// TIA Portal V20 export
FUNCTION_BLOCK "CONTROL_LINE"   // FB7, LAD
{ S7_Optimized_Access := 'TRUE' }
// stored: MemoryReserve 100, SetENOAutomatically false
   VAR
      TIMER_reset { S7_SetPoint := 'True'} : TON_TIME;
      P_TRIG_INICIAL : Bool;
      P_TRIG_RESET : Bool;
      AUTOMAT { S7_SetPoint := 'True'} : "SENSOR";
      MANUAL { S7_SetPoint := 'True'} : "SENSOR";
      SENSOR_3 { S7_SetPoint := 'True'} : "SENSOR";
      SENSOR_4 { S7_SetPoint := 'True'} : "SENSOR";
      SENSOR_5 { S7_SetPoint := 'True'} : "SENSOR";
      SENSOR_6 { S7_SetPoint := 'True'} : "SENSOR";
      SENSOR_7 { S7_SetPoint := 'True'} : "SENSOR";
      SENSOR_8 { S7_SetPoint := 'True'} : "SENSOR";
      SENSOR_9 { S7_SetPoint := 'True'} : "SENSOR";
      SENSOR_10 { S7_SetPoint := 'True'} : "SENSOR";
      SENSOR_11 { S7_SetPoint := 'True'} : "SENSOR";
      dvere_L_A { S7_SetPoint := 'True'} : "SENSOR";
      dvere_L_B { S7_SetPoint := 'True'} : "SENSOR";
      dvere_P_A { S7_SetPoint := 'True'} : "SENSOR";
      dvere_P_B { S7_SetPoint := 'True'} : "SENSOR";
      SEN_STRUCT : Struct
         AUTOMAT : Bool;
         AUTOMAT_NEG : Bool;
         MANUAL : Bool;
         MANUAL_NEG : Bool;
         SENSOR_TLAKU : Bool;
         SENSOR_TLAKU_NEG : Bool;
         power : Bool;
         power_neg : Bool;
         safety : Bool;
         safety_neg : Bool;
         s_10 : Bool;
         TLA_STOP : Bool;
         TLA_STOP_NEG : Bool;
         TLA_START : Bool;
         TLA_START_NEG : Bool;
         TLA_KVIT : Bool;
         TLA_KVIT_NEG : Bool;
         s_17 : Bool;
         S19 : Bool;
         L1_OK : Bool;
         L1_NOT_OK : Bool;
         L2_OK : Bool;
         L2_NOT_OK : Bool;
         L3_OK : Bool;
         L3_NOT_OK : Bool;
         dvere_L_A : Bool;
         dvere_L_B : Bool;
         dvere_P_A : Bool;
         dvere_P_B : Bool;
         S30 : Bool;
         S31 : Bool;
         LASER_MEMOR : Bool;
      END_STRUCT;
      "M" : Struct
         P_TRIK_hmi_manual : Bool;
         p_trig_hmi_automat : Bool;
         N_TRIG_REZIM : Bool;
         M_4 : Bool;
         hlaseni_chyby : Bool;
         M_6 : Bool;
         M_7 : Bool;
         M_8 : Bool;
         M_9 : Bool;
         p_Trig_al : Bool;
         n_trig_al : Bool;
         p_trig_wro : Bool;
         n_trig_wro : Bool;
         M_14 : Bool;
         M_15 : Bool;
         N_TRIG_MANUAL : Bool;
         M_17 : Bool;
         M_18 : Bool;
         M_19 : Bool;
         M_20 : Bool;
         M_21 : Bool;
         M_22 : Bool;
         M_23 : Bool;
         M_24 : Bool;
         M_25 : Bool;
         M_26 : Bool;
         M_27 : Bool;
         M_28 : Bool;
         M_29 : Bool;
         M_30 : Bool;
         M_31 : Bool;
         M_32 : Bool;
      END_STRUCT;
      trig : Struct
         reset_error_all : Bool;
         TRIG_FOR_OP_4_AUTOMAT : Bool;
         t_3 : Bool;
         t_4 : Bool;
         t_5 : Bool;
         t_6 : Bool;
         t_7 : Bool;
         t_8 : Bool;
      END_STRUCT;
      SQCR : Int;
      job_mailbox : Array[0..3] of Word;
      n_trig_res_auit : Bool;
      inicial_control { S7_SetPoint := 'True'} : TON_TIME;
      SQCR_SAFETY { S7_SetPoint := 'True'} : Int;
      n_trig_RESET_AUT : Bool;
      P_TRIG_RESET_SAFETY : Bool;
      air { S7_SetPoint := 'True'} : TON_TIME;
      HMI_ALARM { S7_SetPoint := 'True'} : Int;
   END_VAR
   VAR_TEMP
      "string" : String;
      smaz_me : Bool;
      majak_green_s1 : Bool;
      majak_red_s1 : Bool;
      majak_yelou_s1 : Bool;
      majak_blue_s1 : Bool;
      majak_orange_s1 : Bool;
      majak_green_s2 : Bool;
      majak_red_s2 : Bool;
      majak_yelou_s2 : Bool;
      majak_blue_s2 : Bool;
      majak_orange_s2 : Bool;
      majak_green_s3 : Bool;
      majak_red_s3 : Bool;
      majak_yelou_s3 : Bool;
      majak_blue_s3 : Bool;
      majak_orange_s3 : Bool;
      majak_green_s4 : Bool;
      majak_red_s4 : Bool;
      majak_yelou_s4 : Bool;
      majak_blue_s4 : Bool;
      majak_orange_s4 : Bool;
      majak_green_s5 : Bool;
      majak_red_s5 : Bool;
      majak_yelou_s5 : Bool;
      majak_blue_s5 : Bool;
      majak_orange_s5 : Bool;
   END_VAR
   VAR CONSTANT
      STEP_0_FIRST_START : Int := 0;
      STEP_3 : Int := 3;
      STEP_5 : Int := 5;
      STEP_10 : Int := 10;
      STEP_15 : Int := 15;
      STEP_20 : Int := 20;
      STEP_25 : Int := 25;
      STEP_27 : Int := 27;
      STEP_30 : Int := 30;
      STEP_35 : Int := 35;
      STEP_40 : Int := 40;
      STEP_45 : Int := 45;
      STEP_48 : Int := 48;
      STEP_50 : Int := 50;
      STEP_52 : Int := 52;
      STEP_55 : Int := 55;
      STEP_60 : Int := 60;
      STEP_65 : Int := 65;
      STEP_70 : Int := 70;
      STEP_75 : Int := 75;
      STEP_80 : Int := 80;
      STEP_85 : Int := 85;
      STEP_90 : Int := 90;
      STEP_95 : Int := 95;
      STEP_100 : Int := 100;
      STEO_105 : Int := 105;
   END_VAR
   VAR_TEMP   // added for the SCL form of the ladder/FBD networks
      _w1 : Bool;
      _w2 : Bool;
      _w3 : Bool;
      _w4 : Bool;
      _w5 : Bool;
   END_VAR
BEGIN

REGION Network 1 (SCL)
   // SET  BASIC ELEMENTS
   // odpojení nepoužívaných kontaktů
   "LOG_0" := 0;
   "LOG_1" := 1;
   "SMAZ_ME_0" := 0;
   "SMAZ_ME_1" := 1;
END_REGION

REGION Network 2: SENSORS
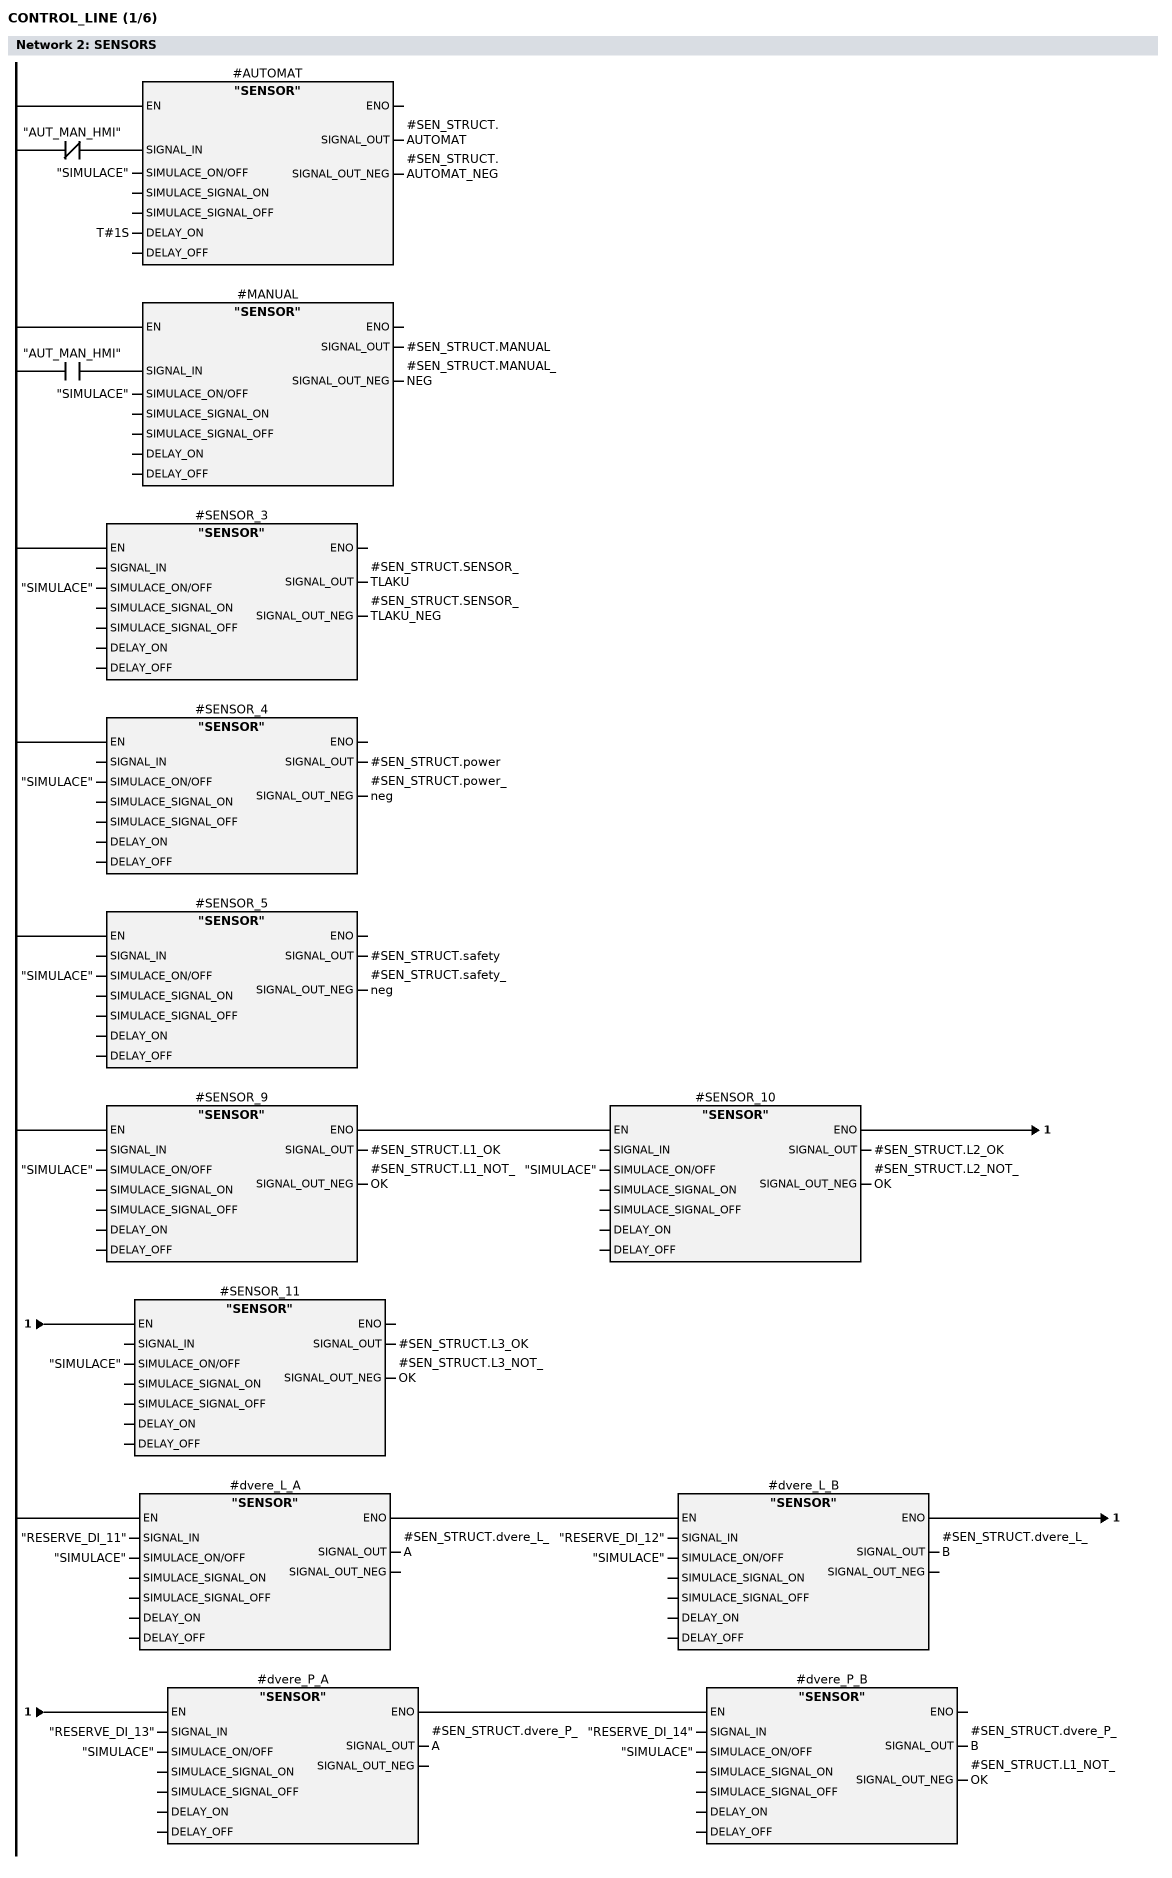
   RUNG wire#powerrail
      #AUTOMAT(SIGNAL_IN := wire#w1, "SIMULACE_ON/OFF" := "SIMULACE", SIMULACE_SIGNAL_ON :=, SIMULACE_SIGNAL_OFF :=, DELAY_ON := T#1S, DELAY_OFF :=, SIGNAL_OUT => #SEN_STRUCT.AUTOMAT, SIGNAL_OUT_NEG => #SEN_STRUCT.AUTOMAT_NEG)
   END_RUNG
   RUNG wire#powerrail
      I_Contact( "AUT_MAN_HMI" )
   END_RUNG wire#w1
   RUNG wire#powerrail
      #MANUAL(SIGNAL_IN := wire#w2, "SIMULACE_ON/OFF" := "SIMULACE", SIMULACE_SIGNAL_ON :=, SIMULACE_SIGNAL_OFF :=, DELAY_ON :=, DELAY_OFF :=, SIGNAL_OUT => #SEN_STRUCT.MANUAL, SIGNAL_OUT_NEG => #SEN_STRUCT.MANUAL_NEG)
   END_RUNG
   RUNG wire#powerrail
      Contact( "AUT_MAN_HMI" )
   END_RUNG wire#w2
   RUNG wire#powerrail
      #SENSOR_3(SIGNAL_IN :=, "SIMULACE_ON/OFF" := "SIMULACE", SIMULACE_SIGNAL_ON :=, SIMULACE_SIGNAL_OFF :=, DELAY_ON :=, DELAY_OFF :=, SIGNAL_OUT => #SEN_STRUCT.SENSOR_TLAKU, SIGNAL_OUT_NEG => #SEN_STRUCT.SENSOR_TLAKU_NEG)
   END_RUNG
   RUNG wire#powerrail
      #SENSOR_4(SIGNAL_IN :=, "SIMULACE_ON/OFF" := "SIMULACE", SIMULACE_SIGNAL_ON :=, SIMULACE_SIGNAL_OFF :=, DELAY_ON :=, DELAY_OFF :=, SIGNAL_OUT => #SEN_STRUCT.power, SIGNAL_OUT_NEG => #SEN_STRUCT.power_neg)
   END_RUNG
   RUNG wire#powerrail
      #SENSOR_5(SIGNAL_IN :=, "SIMULACE_ON/OFF" := "SIMULACE", SIMULACE_SIGNAL_ON :=, SIMULACE_SIGNAL_OFF :=, DELAY_ON :=, DELAY_OFF :=, SIGNAL_OUT => #SEN_STRUCT.safety, SIGNAL_OUT_NEG => #SEN_STRUCT.safety_neg)
   END_RUNG
   RUNG wire#powerrail
      #SENSOR_9(SIGNAL_IN :=, "SIMULACE_ON/OFF" := "SIMULACE", SIMULACE_SIGNAL_ON :=, SIMULACE_SIGNAL_OFF :=, DELAY_ON :=, DELAY_OFF :=, SIGNAL_OUT => #SEN_STRUCT.L1_OK, SIGNAL_OUT_NEG => #SEN_STRUCT.L1_NOT_OK)
      #SENSOR_10(SIGNAL_IN :=, "SIMULACE_ON/OFF" := "SIMULACE", SIMULACE_SIGNAL_ON :=, SIMULACE_SIGNAL_OFF :=, DELAY_ON :=, DELAY_OFF :=, SIGNAL_OUT => #SEN_STRUCT.L2_OK, SIGNAL_OUT_NEG => #SEN_STRUCT.L2_NOT_OK)
      #SENSOR_11(SIGNAL_IN :=, "SIMULACE_ON/OFF" := "SIMULACE", SIMULACE_SIGNAL_ON :=, SIMULACE_SIGNAL_OFF :=, DELAY_ON :=, DELAY_OFF :=, SIGNAL_OUT => #SEN_STRUCT.L3_OK, SIGNAL_OUT_NEG => #SEN_STRUCT.L3_NOT_OK)
   END_RUNG
   RUNG wire#powerrail
      #dvere_L_A(SIGNAL_IN := "RESERVE_DI_11", "SIMULACE_ON/OFF" := "SIMULACE", SIMULACE_SIGNAL_ON :=, SIMULACE_SIGNAL_OFF :=, DELAY_ON :=, DELAY_OFF :=, SIGNAL_OUT => #SEN_STRUCT.dvere_L_A, SIGNAL_OUT_NEG =>)
      #dvere_L_B(SIGNAL_IN := "RESERVE_DI_12", "SIMULACE_ON/OFF" := "SIMULACE", SIMULACE_SIGNAL_ON :=, SIMULACE_SIGNAL_OFF :=, DELAY_ON :=, DELAY_OFF :=, SIGNAL_OUT => #SEN_STRUCT.dvere_L_B, SIGNAL_OUT_NEG =>)
      #dvere_P_A(SIGNAL_IN := "RESERVE_DI_13", "SIMULACE_ON/OFF" := "SIMULACE", SIMULACE_SIGNAL_ON :=, SIMULACE_SIGNAL_OFF :=, DELAY_ON :=, DELAY_OFF :=, SIGNAL_OUT => #SEN_STRUCT.dvere_P_A, SIGNAL_OUT_NEG =>)
      #dvere_P_B(SIGNAL_IN := "RESERVE_DI_14", "SIMULACE_ON/OFF" := "SIMULACE", SIMULACE_SIGNAL_ON :=, SIMULACE_SIGNAL_OFF :=, DELAY_ON :=, DELAY_OFF :=, SIGNAL_OUT => #SEN_STRUCT.dvere_P_B, SIGNAL_OUT_NEG => #SEN_STRUCT.L1_NOT_OK)
   END_RUNG
   // the same network as SCL:
   #AUTOMAT(SIGNAL_IN := NOT "AUT_MAN_HMI",   // "SENSOR"
            "SIMULACE_ON/OFF" := "SIMULACE",
            DELAY_ON := T#1S,
            SIGNAL_OUT => #SEN_STRUCT.AUTOMAT,
            SIGNAL_OUT_NEG => #SEN_STRUCT.AUTOMAT_NEG);
   #MANUAL(SIGNAL_IN := "AUT_MAN_HMI",   // "SENSOR"
           "SIMULACE_ON/OFF" := "SIMULACE",
           SIGNAL_OUT => #SEN_STRUCT.MANUAL,
           SIGNAL_OUT_NEG => #SEN_STRUCT.MANUAL_NEG);
   #SENSOR_3("SIMULACE_ON/OFF" := "SIMULACE",   // "SENSOR"
             SIGNAL_OUT => #SEN_STRUCT.SENSOR_TLAKU,
             SIGNAL_OUT_NEG => #SEN_STRUCT.SENSOR_TLAKU_NEG);
   #SENSOR_4("SIMULACE_ON/OFF" := "SIMULACE",   // "SENSOR"
             SIGNAL_OUT => #SEN_STRUCT.power,
             SIGNAL_OUT_NEG => #SEN_STRUCT.power_neg);
   #SENSOR_5("SIMULACE_ON/OFF" := "SIMULACE",   // "SENSOR"
             SIGNAL_OUT => #SEN_STRUCT.safety,
             SIGNAL_OUT_NEG => #SEN_STRUCT.safety_neg);
   #SENSOR_9("SIMULACE_ON/OFF" := "SIMULACE",   // "SENSOR"
             SIGNAL_OUT => #SEN_STRUCT.L1_OK,
             SIGNAL_OUT_NEG => #SEN_STRUCT.L1_NOT_OK,
             ENO => #_w1);
   #SENSOR_10(EN := #_w1,   // "SENSOR"
              "SIMULACE_ON/OFF" := "SIMULACE",
              SIGNAL_OUT => #SEN_STRUCT.L2_OK,
              SIGNAL_OUT_NEG => #SEN_STRUCT.L2_NOT_OK,
              ENO => #_w2);
   IF #_w2 THEN
       #SENSOR_11("SIMULACE_ON/OFF" := "SIMULACE",   // "SENSOR"
                  SIGNAL_OUT => #SEN_STRUCT.L3_OK,
                  SIGNAL_OUT_NEG => #SEN_STRUCT.L3_NOT_OK);
   END_IF;
   #dvere_L_A(SIGNAL_IN := "RESERVE_DI_11",   // "SENSOR"
              "SIMULACE_ON/OFF" := "SIMULACE",
              SIGNAL_OUT => #SEN_STRUCT.dvere_L_A,
              ENO => #_w3);
   #dvere_L_B(EN := #_w3,   // "SENSOR"
              SIGNAL_IN := "RESERVE_DI_12",
              "SIMULACE_ON/OFF" := "SIMULACE",
              SIGNAL_OUT => #SEN_STRUCT.dvere_L_B,
              ENO => #_w4);
   #dvere_P_A(EN := #_w4,   // "SENSOR"
              SIGNAL_IN := "RESERVE_DI_13",
              "SIMULACE_ON/OFF" := "SIMULACE",
              SIGNAL_OUT => #SEN_STRUCT.dvere_P_A,
              ENO => #_w5);
   IF #_w5 THEN
       #dvere_P_B(SIGNAL_IN := "RESERVE_DI_14",   // "SENSOR"
                  "SIMULACE_ON/OFF" := "SIMULACE",
                  SIGNAL_OUT => #SEN_STRUCT.dvere_P_B,
                  SIGNAL_OUT_NEG => #SEN_STRUCT.L1_NOT_OK);
   END_IF;
END_REGION

REGION Network 3 (SCL): ALARMY OP1/OP2 -> HMI
   // ===== ALARMY -> HMI (DB_ALARM.alarm_line, HMI ID 1-16) =====
   // bit 9 (ID 10 aplikator) a bit 14 (ID 15 tlak vzduchu) = firemni standard, nepouzivat

   // bit 0 - tiskarna nekomunikuje (OP2 se nevrati do kroku 5 do 15 s)
   "DB_ALARM".T_tiskarna.TON(IN := "AUTOMAT" AND "OP2_DB".SQCR <> 5,
                             PT := T#15S);
   "DB_ALARM".alarm_line.%X0 := "DB_ALARM".T_tiskarna.Q;

   // bity 1-3 - kamery offline (jen v automatu)
   "DB_ALARM".alarm_line.%X1 := "AUTOMAT" AND NOT "COG_FOLIE_L_is3800-Online";
   "DB_ALARM".alarm_line.%X2 := "AUTOMAT" AND NOT "COG_FOLIE_P_is3800-Online";
   "DB_ALARM".alarm_line.%X3 := "AUTOMAT" AND NOT "COG_ETIKETA_is3800-Online"
   AND NOT "OP1_DB".Kam_Etiketa_Job.aktivni;   // pri loadu jobu je kamera chvili offline

   // bit 4 - chybne datum v recepture
   "DB_ALARM".alarm_line.%X4 := "OP2_DB".Tisk.datum_chyba;

   // bit 5 - fronta plna
   "DB_ALARM".alarm_line.%X5 := "OP1_DB".Kamera.fronta_plna;

   // bit 6 - job horni kamery se nenacetl
   //"DB_ALARM".alarm_line.%X6 := "OP1_DB".Kam_Etiketa_Job.chyba;

   // bity 7-8 - otevrene dvere (signaly ze site "alarmy")
   "DB_ALARM".alarm_line.%X7 := "DB_ALARM".WRONG.dvere_L_tevreny;
   "DB_ALARM".alarm_line.%X8 := "DB_ALARM".WRONG.dvere_P_otevreny;

   // souhrnny alarm -> KA19 blika, HMI_ALARM = 10
   "alrm_global" := "DB_ALARM".alarm_line <> 0;
   "DB_ALARM".ALARM.ALARM_GLOBAL := "alrm_global";
END_REGION

REGION Network 4: alarmy
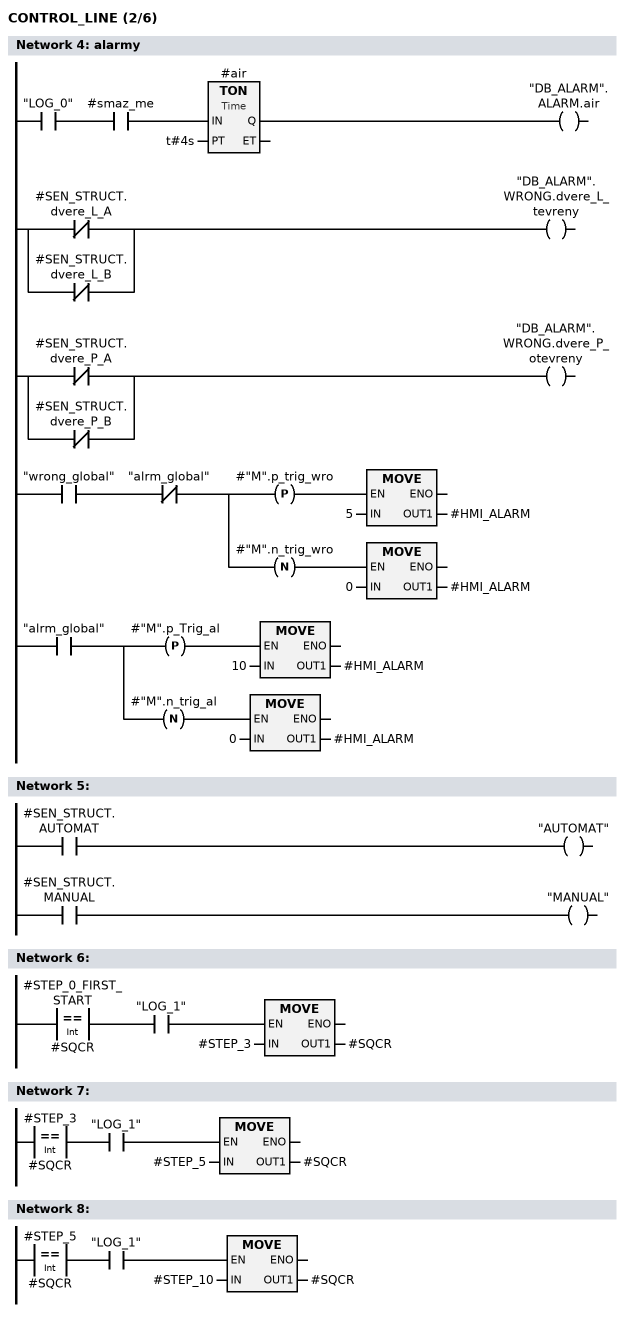
   RUNG wire#powerrail
      Contact( "LOG_0" )
      Contact( #smaz_me )
      { S7_Templates := "time_type := Time" } #air.TON(pt := t#4s, et =>)
      Coil( "DB_ALARM".ALARM.air )
   END_RUNG
   RUNG wire#powerrail
      I_Contact( #SEN_STRUCT.dvere_L_A )
      wire#w1
      Coil( "DB_ALARM".WRONG.dvere_L_tevreny )
   END_RUNG
   RUNG wire#powerrail
      I_Contact( #SEN_STRUCT.dvere_L_B )
   END_RUNG wire#w1
   RUNG wire#powerrail
      I_Contact( #SEN_STRUCT.dvere_P_A )
      wire#w2
      Coil( "DB_ALARM".WRONG.dvere_P_otevreny )
   END_RUNG
   RUNG wire#powerrail
      I_Contact( #SEN_STRUCT.dvere_P_B )
   END_RUNG wire#w2
   RUNG wire#powerrail
      Contact( "wrong_global" )
      I_Contact( "alrm_global" )
      wire#w3
      P_Trig( #"M".p_trig_wro )
      Move(in := 5, out1 => #HMI_ALARM)
   END_RUNG
   RUNG wire#w3
      N_Trig( #"M".n_trig_wro )
      Move(in := 0, out1 => #HMI_ALARM)
   END_RUNG
   RUNG wire#powerrail
      Contact( "alrm_global" )
      wire#w4
      P_Trig( #"M".p_Trig_al )
      Move(in := 10, out1 => #HMI_ALARM)
   END_RUNG
   RUNG wire#w4
      N_Trig( #"M".n_trig_al )
      Move(in := 0, out1 => #HMI_ALARM)
   END_RUNG
   // the same network as SCL:
   #air(IN := "LOG_0" AND #smaz_me, PT := t#4s);   // TON
   "DB_ALARM".ALARM.air := #air.Q;
   "DB_ALARM".WRONG.dvere_L_tevreny := NOT #SEN_STRUCT.dvere_L_A OR NOT #SEN_STRUCT.dvere_L_B;
   "DB_ALARM".WRONG.dvere_P_otevreny := NOT #SEN_STRUCT.dvere_P_A OR NOT #SEN_STRUCT.dvere_P_B;
   #_w1 := "wrong_global" AND NOT "alrm_global";
   #_w2 := #_w1 AND NOT #"M".p_trig_wro;   // rising edge
   #"M".p_trig_wro := #_w1;
   IF #_w2 THEN #HMI_ALARM := 5; END_IF;
   #_w3 := NOT #_w1 AND #"M".n_trig_wro;   // falling edge
   #"M".n_trig_wro := #_w1;
   IF #_w3 THEN #HMI_ALARM := 0; END_IF;
   #_w4 := "alrm_global" AND NOT #"M".p_Trig_al;   // rising edge
   #"M".p_Trig_al := "alrm_global";
   IF #_w4 THEN #HMI_ALARM := 10; END_IF;
   #_w5 := NOT "alrm_global" AND #"M".n_trig_al;   // falling edge
   #"M".n_trig_al := "alrm_global";
   IF #_w5 THEN #HMI_ALARM := 0; END_IF;
END_REGION

REGION Network 5
   RUNG wire#powerrail
      Contact( #SEN_STRUCT.AUTOMAT )
      Coil( "AUTOMAT" )
   END_RUNG
   RUNG wire#powerrail
      Contact( #SEN_STRUCT.MANUAL )
      Coil( "MANUAL" )
   END_RUNG
   // the same network as SCL:
   "AUTOMAT" := #SEN_STRUCT.AUTOMAT;
   "MANUAL" := #SEN_STRUCT.MANUAL;
END_REGION

REGION Network 6
   RUNG wire#powerrail
      { S7_Templates := "SrcType := Int" } EQ_Contact(in1 := #STEP_0_FIRST_START, in2 := #SQCR)
      Contact( "LOG_1" )
      Move(in := #STEP_3, out1 => #SQCR)
   END_RUNG
   // the same network as SCL:
   IF (#STEP_0_FIRST_START = #SQCR) AND "LOG_1" THEN #SQCR := #STEP_3; END_IF;
END_REGION

REGION Network 7
   RUNG wire#powerrail
      { S7_Templates := "SrcType := Int" } EQ_Contact(in1 := #STEP_3, in2 := #SQCR)
      Contact( "LOG_1" )
      Move(in := #STEP_5, out1 => #SQCR)
   END_RUNG
   // the same network as SCL:
   IF (#STEP_3 = #SQCR) AND "LOG_1" THEN #SQCR := #STEP_5; END_IF;
END_REGION

REGION Network 8
   RUNG wire#powerrail
      { S7_Templates := "SrcType := Int" } EQ_Contact(in1 := #STEP_5, in2 := #SQCR)
      Contact( "LOG_1" )
      Move(in := #STEP_10, out1 => #SQCR)
   END_RUNG
   // the same network as SCL:
   IF (#STEP_5 = #SQCR) AND "LOG_1" THEN #SQCR := #STEP_10; END_IF;
END_REGION

REGION Network 9
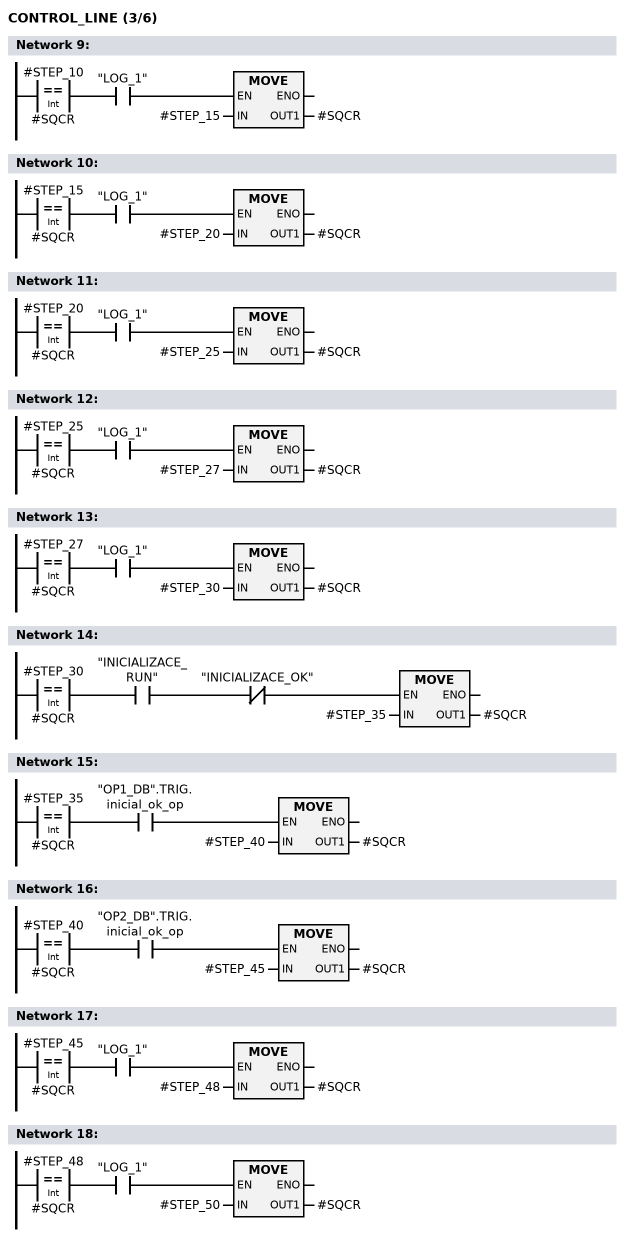
   RUNG wire#powerrail
      { S7_Templates := "SrcType := Int" } EQ_Contact(in1 := #STEP_10, in2 := #SQCR)
      Contact( "LOG_1" )
      Move(in := #STEP_15, out1 => #SQCR)
   END_RUNG
   // the same network as SCL:
   IF (#STEP_10 = #SQCR) AND "LOG_1" THEN #SQCR := #STEP_15; END_IF;
END_REGION

REGION Network 10
   RUNG wire#powerrail
      { S7_Templates := "SrcType := Int" } EQ_Contact(in1 := #STEP_15, in2 := #SQCR)
      Contact( "LOG_1" )
      Move(in := #STEP_20, out1 => #SQCR)
   END_RUNG
   // the same network as SCL:
   IF (#STEP_15 = #SQCR) AND "LOG_1" THEN #SQCR := #STEP_20; END_IF;
END_REGION

REGION Network 11
   RUNG wire#powerrail
      { S7_Templates := "SrcType := Int" } EQ_Contact(in1 := #STEP_20, in2 := #SQCR)
      Contact( "LOG_1" )
      Move(in := #STEP_25, out1 => #SQCR)
   END_RUNG
   // the same network as SCL:
   IF (#STEP_20 = #SQCR) AND "LOG_1" THEN #SQCR := #STEP_25; END_IF;
END_REGION

REGION Network 12
   RUNG wire#powerrail
      { S7_Templates := "SrcType := Int" } EQ_Contact(in1 := #STEP_25, in2 := #SQCR)
      Contact( "LOG_1" )
      Move(in := #STEP_27, out1 => #SQCR)
   END_RUNG
   // the same network as SCL:
   IF (#STEP_25 = #SQCR) AND "LOG_1" THEN #SQCR := #STEP_27; END_IF;
END_REGION

REGION Network 13
   RUNG wire#powerrail
      { S7_Templates := "SrcType := Int" } EQ_Contact(in1 := #STEP_27, in2 := #SQCR)
      Contact( "LOG_1" )
      Move(in := #STEP_30, out1 => #SQCR)
   END_RUNG
   // the same network as SCL:
   IF (#STEP_27 = #SQCR) AND "LOG_1" THEN #SQCR := #STEP_30; END_IF;
END_REGION

REGION Network 14
   RUNG wire#powerrail
      { S7_Templates := "SrcType := Int" } EQ_Contact(in1 := #STEP_30, in2 := #SQCR)
      Contact( "INICIALIZACE_RUN" )
      I_Contact( "INICIALIZACE_OK" )
      Move(in := #STEP_35, out1 => #SQCR)
   END_RUNG
   // the same network as SCL:
   IF (#STEP_30 = #SQCR) AND "INICIALIZACE_RUN" AND NOT "INICIALIZACE_OK" THEN #SQCR := #STEP_35; END_IF;
END_REGION

REGION Network 15
   RUNG wire#powerrail
      { S7_Templates := "SrcType := Int" } EQ_Contact(in1 := #STEP_35, in2 := #SQCR)
      Contact( "OP1_DB".TRIG.inicial_ok_op )
      Move(in := #STEP_40, out1 => #SQCR)
   END_RUNG
   // the same network as SCL:
   IF (#STEP_35 = #SQCR) AND "OP1_DB".TRIG.inicial_ok_op THEN #SQCR := #STEP_40; END_IF;
END_REGION

REGION Network 16
   RUNG wire#powerrail
      { S7_Templates := "SrcType := Int" } EQ_Contact(in1 := #STEP_40, in2 := #SQCR)
      Contact( "OP2_DB".TRIG.inicial_ok_op )
      Move(in := #STEP_45, out1 => #SQCR)
   END_RUNG
   // the same network as SCL:
   IF (#STEP_40 = #SQCR) AND "OP2_DB".TRIG.inicial_ok_op THEN #SQCR := #STEP_45; END_IF;
END_REGION

REGION Network 17
   RUNG wire#powerrail
      { S7_Templates := "SrcType := Int" } EQ_Contact(in1 := #STEP_45, in2 := #SQCR)
      Contact( "LOG_1" )
      Move(in := #STEP_48, out1 => #SQCR)
   END_RUNG
   // the same network as SCL:
   IF (#STEP_45 = #SQCR) AND "LOG_1" THEN #SQCR := #STEP_48; END_IF;
END_REGION

REGION Network 18
   RUNG wire#powerrail
      { S7_Templates := "SrcType := Int" } EQ_Contact(in1 := #STEP_48, in2 := #SQCR)
      Contact( "LOG_1" )
      Move(in := #STEP_50, out1 => #SQCR)
   END_RUNG
   // the same network as SCL:
   IF (#STEP_48 = #SQCR) AND "LOG_1" THEN #SQCR := #STEP_50; END_IF;
END_REGION

REGION Network 19
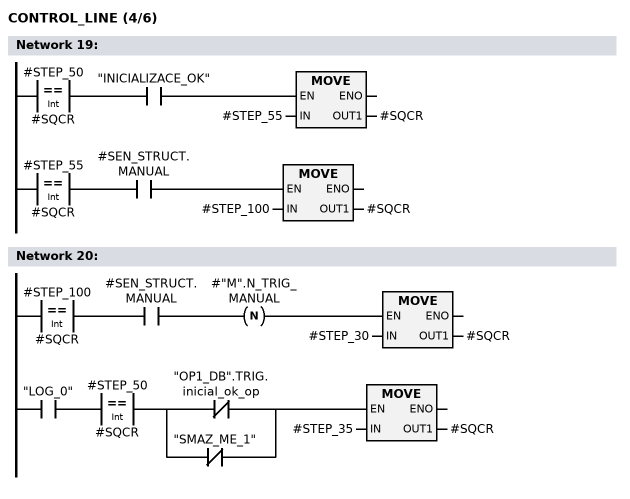
   RUNG wire#powerrail
      { S7_Templates := "SrcType := Int" } EQ_Contact(in1 := #STEP_50, in2 := #SQCR)
      Contact( "INICIALIZACE_OK" )
      Move(in := #STEP_55, out1 => #SQCR)
   END_RUNG
   RUNG wire#powerrail
      { S7_Templates := "SrcType := Int" } EQ_Contact(in1 := #STEP_55, in2 := #SQCR)
      Contact( #SEN_STRUCT.MANUAL )
      Move(in := #STEP_100, out1 => #SQCR)
   END_RUNG
   // the same network as SCL:
   IF (#STEP_50 = #SQCR) AND "INICIALIZACE_OK" THEN #SQCR := #STEP_55; END_IF;
   IF (#STEP_55 = #SQCR) AND #SEN_STRUCT.MANUAL THEN #SQCR := #STEP_100; END_IF;
END_REGION

REGION Network 20
   RUNG wire#powerrail
      { S7_Templates := "SrcType := Int" } EQ_Contact(in1 := #STEP_100, in2 := #SQCR)
      Contact( #SEN_STRUCT.MANUAL )
      N_Trig( #"M".N_TRIG_MANUAL )
      Move(in := #STEP_30, out1 => #SQCR)
   END_RUNG
   RUNG wire#powerrail
      Contact( "LOG_0" )
      { S7_Templates := "SrcType := Int" } EQ_Contact(in1 := #STEP_50, in2 := #SQCR)
      wire#w1
      I_Contact( "OP1_DB".TRIG.inicial_ok_op )
      wire#w2
      Move(in := #STEP_35, out1 => #SQCR)
   END_RUNG
   RUNG wire#w1
      I_Contact( "SMAZ_ME_1" )
   END_RUNG wire#w2
   // the same network as SCL:
   #_w1 := (#STEP_100 = #SQCR) AND #SEN_STRUCT.MANUAL;
   #_w2 := NOT #_w1 AND #"M".N_TRIG_MANUAL;   // falling edge
   #"M".N_TRIG_MANUAL := #_w1;
   IF #_w2 THEN #SQCR := #STEP_30; END_IF;
   IF "LOG_0" AND (#STEP_50 = #SQCR) AND (NOT "OP1_DB".TRIG.inicial_ok_op OR NOT "SMAZ_ME_1") THEN
       #SQCR := #STEP_35;
   END_IF;
END_REGION

REGION Network 21: LEDKY
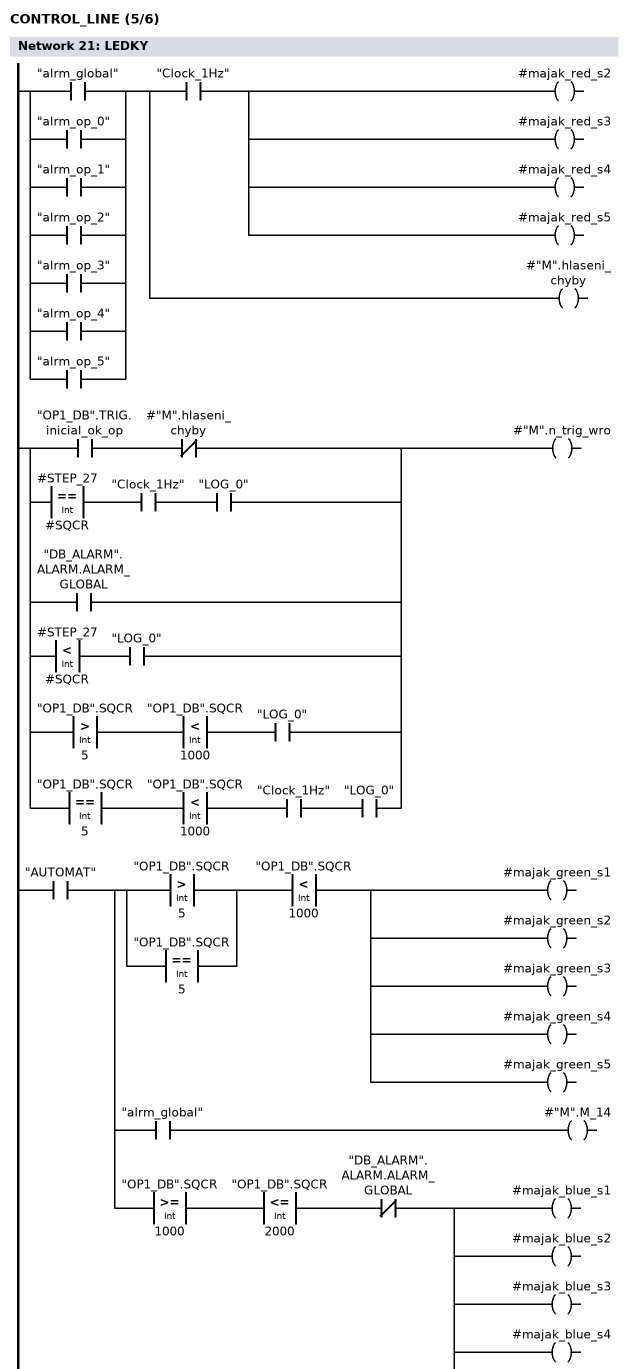
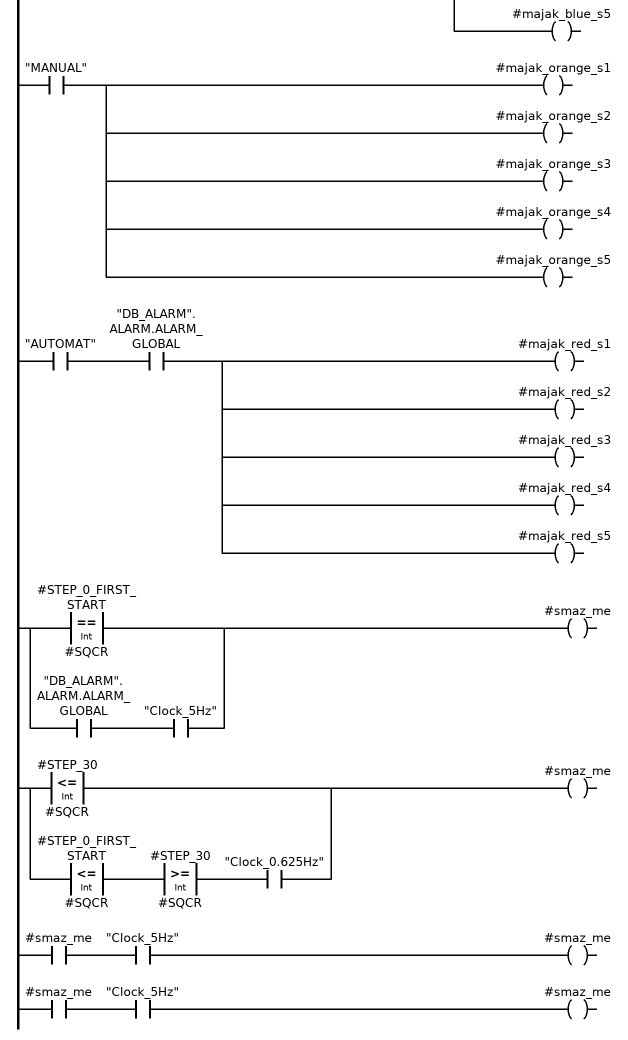
   RUNG wire#powerrail
      Contact( "alrm_global" )
      wire#w1
      Contact( "Clock_1Hz" )
      wire#w2
      Coil( #majak_red_s2 )
   END_RUNG
   RUNG wire#powerrail
      Contact( "alrm_op_0" )
   END_RUNG wire#w1
   RUNG wire#powerrail
      Contact( "alrm_op_1" )
   END_RUNG wire#w1
   RUNG wire#powerrail
      Contact( "alrm_op_2" )
   END_RUNG wire#w1
   RUNG wire#powerrail
      Contact( "alrm_op_3" )
   END_RUNG wire#w1
   RUNG wire#powerrail
      Contact( "alrm_op_4" )
   END_RUNG wire#w1
   RUNG wire#powerrail
      Contact( "alrm_op_5" )
   END_RUNG wire#w1
   RUNG wire#w2
      Coil( #majak_red_s3 )
   END_RUNG
   RUNG wire#w2
      Coil( #majak_red_s4 )
   END_RUNG
   RUNG wire#w2
      Coil( #majak_red_s5 )
   END_RUNG
   RUNG wire#w1
      Coil( #"M".hlaseni_chyby )
   END_RUNG
   RUNG wire#powerrail
      Contact( "OP1_DB".TRIG.inicial_ok_op )
      I_Contact( #"M".hlaseni_chyby )
      wire#w3
      Coil( #"M".n_trig_wro )
   END_RUNG
   RUNG wire#powerrail
      { S7_Templates := "SrcType := Int" } EQ_Contact(in1 := #STEP_27, in2 := #SQCR)
      Contact( "Clock_1Hz" )
      Contact( "LOG_0" )
   END_RUNG wire#w3
   RUNG wire#powerrail
      Contact( "DB_ALARM".ALARM.ALARM_GLOBAL )
   END_RUNG wire#w3
   RUNG wire#powerrail
      { S7_Templates := "SrcType := Int" } LT_Contact(in1 := #STEP_27, in2 := #SQCR)
      Contact( "LOG_0" )
   END_RUNG wire#w3
   RUNG wire#powerrail
      { S7_Templates := "SrcType := Int" } GT_Contact(in1 := "OP1_DB".SQCR, in2 := 5)
      { S7_Templates := "SrcType := Int" } LT_Contact(in1 := "OP1_DB".SQCR, in2 := 1000)
      Contact( "LOG_0" )
   END_RUNG wire#w3
   RUNG wire#powerrail
      { S7_Templates := "SrcType := Int" } EQ_Contact(in1 := "OP1_DB".SQCR, in2 := 5)
      { S7_Templates := "SrcType := Int" } LT_Contact(in1 := "OP1_DB".SQCR, in2 := 1000)
      Contact( "Clock_1Hz" )
      Contact( "LOG_0" )
   END_RUNG wire#w3
   RUNG wire#powerrail
      Contact( "AUTOMAT" )
      wire#w4
      { S7_Templates := "SrcType := Int" } GT_Contact(in1 := "OP1_DB".SQCR, in2 := 5)
      wire#w5
      { S7_Templates := "SrcType := Int" } LT_Contact(in1 := "OP1_DB".SQCR, in2 := 1000)
      wire#w6
      Coil( #majak_green_s1 )
   END_RUNG
   RUNG wire#w4
      { S7_Templates := "SrcType := Int" } EQ_Contact(in1 := "OP1_DB".SQCR, in2 := 5)
   END_RUNG wire#w5
   RUNG wire#w6
      Coil( #majak_green_s2 )
   END_RUNG
   RUNG wire#w6
      Coil( #majak_green_s3 )
   END_RUNG
   RUNG wire#w6
      Coil( #majak_green_s4 )
   END_RUNG
   RUNG wire#w6
      Coil( #majak_green_s5 )
   END_RUNG
   RUNG wire#w4
      Contact( "alrm_global" )
      Coil( #"M".M_14 )
   END_RUNG
   RUNG wire#w4
      { S7_Templates := "SrcType := Int" } GE_Contact(in1 := "OP1_DB".SQCR, in2 := 1000)
      { S7_Templates := "SrcType := Int" } LE_Contact(in1 := "OP1_DB".SQCR, in2 := 2000)
      I_Contact( "DB_ALARM".ALARM.ALARM_GLOBAL )
      wire#w7
      Coil( #majak_blue_s1 )
   END_RUNG
   RUNG wire#w7
      Coil( #majak_blue_s2 )
   END_RUNG
   RUNG wire#w7
      Coil( #majak_blue_s3 )
   END_RUNG
   RUNG wire#w7
      Coil( #majak_blue_s4 )
   END_RUNG
   RUNG wire#w7
      Coil( #majak_blue_s5 )
   END_RUNG
   RUNG wire#powerrail
      Contact( "MANUAL" )
      wire#w8
      Coil( #majak_orange_s1 )
   END_RUNG
   RUNG wire#w8
      Coil( #majak_orange_s2 )
   END_RUNG
   RUNG wire#w8
      Coil( #majak_orange_s3 )
   END_RUNG
   RUNG wire#w8
      Coil( #majak_orange_s4 )
   END_RUNG
   RUNG wire#w8
      Coil( #majak_orange_s5 )
   END_RUNG
   RUNG wire#powerrail
      Contact( "AUTOMAT" )
      Contact( "DB_ALARM".ALARM.ALARM_GLOBAL )
      wire#w9
      Coil( #majak_red_s1 )
   END_RUNG
   RUNG wire#w9
      Coil( #majak_red_s2 )
   END_RUNG
   RUNG wire#w9
      Coil( #majak_red_s3 )
   END_RUNG
   RUNG wire#w9
      Coil( #majak_red_s4 )
   END_RUNG
   RUNG wire#w9
      Coil( #majak_red_s5 )
   END_RUNG
   RUNG wire#powerrail
      { S7_Templates := "SrcType := Int" } EQ_Contact(in1 := #STEP_0_FIRST_START, in2 := #SQCR)
      wire#w10
      Coil( #smaz_me )
   END_RUNG
   RUNG wire#powerrail
      Contact( "DB_ALARM".ALARM.ALARM_GLOBAL )
      Contact( "Clock_5Hz" )
   END_RUNG wire#w10
   RUNG wire#powerrail
      { S7_Templates := "SrcType := Int" } LE_Contact(in1 := #STEP_30, in2 := #SQCR)
      wire#w11
      Coil( #smaz_me )
   END_RUNG
   RUNG wire#powerrail
      { S7_Templates := "SrcType := Int" } LE_Contact(in1 := #STEP_0_FIRST_START, in2 := #SQCR)
      { S7_Templates := "SrcType := Int" } GE_Contact(in1 := #STEP_30, in2 := #SQCR)
      Contact( "Clock_0.625Hz" )
   END_RUNG wire#w11
   RUNG wire#powerrail
      Contact( #smaz_me )
      Contact( "Clock_5Hz" )
      Coil( #smaz_me )
   END_RUNG
   RUNG wire#powerrail
      Contact( #smaz_me )
      Contact( "Clock_5Hz" )
      Coil( #smaz_me )
   END_RUNG
   // the same network as SCL:
   #_w1 := "alrm_global" OR "alrm_op_0" OR "alrm_op_1" OR "alrm_op_2" OR "alrm_op_3" OR "alrm_op_4" OR "alrm_op_5";
   #majak_red_s2 := #_w1 AND "Clock_1Hz";
   #majak_red_s3 := #majak_red_s2;
   #majak_red_s4 := #majak_red_s2;
   #majak_red_s5 := #majak_red_s2;
   #"M".hlaseni_chyby := #_w1;
   #"M".n_trig_wro := ("OP1_DB".TRIG.inicial_ok_op AND NOT #"M".hlaseni_chyby) OR ((#STEP_27 = #SQCR) AND "Clock_1Hz" AND "LOG_0") OR "DB_ALARM".ALARM.ALARM_GLOBAL OR ((#STEP_27 < #SQCR) AND "LOG_0") OR (("OP1_DB".SQCR > 5) AND ("OP1_DB".SQCR < 1000) AND "LOG_0") OR (("OP1_DB".SQCR = 5) AND ("OP1_DB".SQCR < 1000) AND "Clock_1Hz" AND "LOG_0");
   #majak_green_s1 := "AUTOMAT" AND (("OP1_DB".SQCR > 5) OR ("OP1_DB".SQCR = 5)) AND ("OP1_DB".SQCR < 1000);
   #majak_green_s2 := #majak_green_s1;
   #majak_green_s3 := #majak_green_s1;
   #majak_green_s4 := #majak_green_s1;
   #majak_green_s5 := #majak_green_s1;
   #"M".M_14 := "AUTOMAT" AND "alrm_global";
   #majak_blue_s1 := "AUTOMAT" AND ("OP1_DB".SQCR >= 1000) AND ("OP1_DB".SQCR <= 2000) AND NOT "DB_ALARM".ALARM.ALARM_GLOBAL;
   #majak_blue_s2 := #majak_blue_s1;
   #majak_blue_s3 := #majak_blue_s1;
   #majak_blue_s4 := #majak_blue_s1;
   #majak_blue_s5 := #majak_blue_s1;
   #majak_orange_s1 := "MANUAL";
   #majak_orange_s2 := "MANUAL";
   #majak_orange_s3 := "MANUAL";
   #majak_orange_s4 := "MANUAL";
   #majak_orange_s5 := "MANUAL";
   #majak_red_s1 := "AUTOMAT" AND "DB_ALARM".ALARM.ALARM_GLOBAL;
   #majak_red_s2 := #majak_red_s1;
   #majak_red_s3 := #majak_red_s1;
   #majak_red_s4 := #majak_red_s1;
   #majak_red_s5 := #majak_red_s1;
   #smaz_me := (#STEP_0_FIRST_START = #SQCR) OR ("DB_ALARM".ALARM.ALARM_GLOBAL AND "Clock_5Hz");
   #smaz_me := (#STEP_30 <= #SQCR) OR ((#STEP_0_FIRST_START <= #SQCR) AND (#STEP_30 >= #SQCR) AND "Clock_0.625Hz");
   #smaz_me := #smaz_me AND "Clock_5Hz";
   #smaz_me := #smaz_me AND "Clock_5Hz";
END_REGION

REGION Network 22: TRIG EXTERNAL
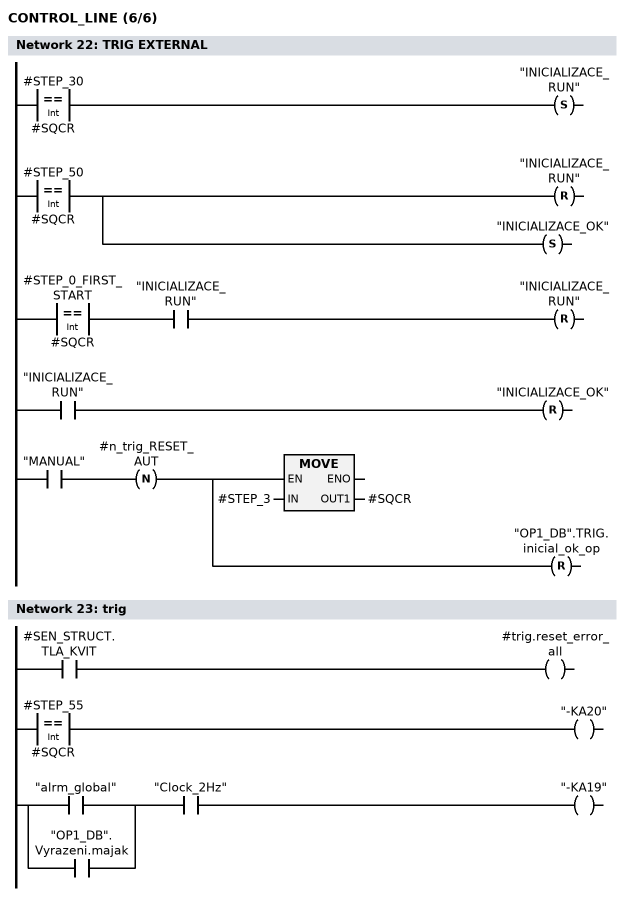
   RUNG wire#powerrail
      { S7_Templates := "SrcType := Int" } EQ_Contact(in1 := #STEP_30, in2 := #SQCR)
      S_Coil( "INICIALIZACE_RUN" )
   END_RUNG
   RUNG wire#powerrail
      { S7_Templates := "SrcType := Int" } EQ_Contact(in1 := #STEP_50, in2 := #SQCR)
      wire#w1
      R_Coil( "INICIALIZACE_RUN" )
   END_RUNG
   RUNG wire#w1
      S_Coil( "INICIALIZACE_OK" )
   END_RUNG
   RUNG wire#powerrail
      { S7_Templates := "SrcType := Int" } EQ_Contact(in1 := #STEP_0_FIRST_START, in2 := #SQCR)
      Contact( "INICIALIZACE_RUN" )
      R_Coil( "INICIALIZACE_RUN" )
   END_RUNG
   RUNG wire#powerrail
      Contact( "INICIALIZACE_RUN" )
      R_Coil( "INICIALIZACE_OK" )
   END_RUNG
   RUNG wire#powerrail
      Contact( "MANUAL" )
      N_Trig( #n_trig_RESET_AUT )
      wire#w2
      Move(in := #STEP_3, out1 => #SQCR)
   END_RUNG
   RUNG wire#w2
      R_Coil( "OP1_DB".TRIG.inicial_ok_op )
   END_RUNG
   // the same network as SCL:
   IF #STEP_30 = #SQCR THEN "INICIALIZACE_RUN" := TRUE; END_IF;
   IF #STEP_50 = #SQCR THEN
       "INICIALIZACE_RUN" := FALSE;
       "INICIALIZACE_OK" := TRUE;
   END_IF;
   IF (#STEP_0_FIRST_START = #SQCR) AND "INICIALIZACE_RUN" THEN "INICIALIZACE_RUN" := FALSE; END_IF;
   IF "INICIALIZACE_RUN" THEN "INICIALIZACE_OK" := FALSE; END_IF;
   #_w1 := NOT "MANUAL" AND #n_trig_RESET_AUT;   // falling edge
   #n_trig_RESET_AUT := "MANUAL";
   IF #_w1 THEN
       #SQCR := #STEP_3;
       "OP1_DB".TRIG.inicial_ok_op := FALSE;
   END_IF;
END_REGION

REGION Network 23: trig
   RUNG wire#powerrail
      Contact( #SEN_STRUCT.TLA_KVIT )
      Coil( #trig.reset_error_all )
   END_RUNG
   RUNG wire#powerrail
      { S7_Templates := "SrcType := Int" } EQ_Contact(in1 := #STEP_55, in2 := #SQCR)
      Coil( "-KA20" )
   END_RUNG
   RUNG wire#powerrail
      Contact( "alrm_global" )
      wire#w1
      Contact( "Clock_2Hz" )
      Coil( "-KA19" )
   END_RUNG
   RUNG wire#powerrail
      Contact( "OP1_DB".Vyrazeni.majak )
   END_RUNG wire#w1
   // the same network as SCL:
   #trig.reset_error_all := #SEN_STRUCT.TLA_KVIT;
   "-KA20" := #STEP_55 = #SQCR;
   "-KA19" := ("alrm_global" OR "OP1_DB".Vyrazeni.majak) AND "Clock_2Hz";
END_REGION
END_FUNCTION_BLOCK
